(* IEC 61131-3 sources: s7-to-codesys/src/POUs/Lang/Converted/FB_ConveyorStl, 2 files *)

(* ---- FB_ConveyorStl.decl.st ---- *)
// Назначение: Конвейер выдачи реагента (STL, таймеры S5)
//             Ленточный конвейер выдачи реагента (STL S7-300); таймеры T1–T5 и счётчик C1 S5 — глобальные.
//             1. Запрос xReq: S по xStart, затем R по xStop OR xJam (сброс главнее; xJam — прошлого вызова).
//             2. Сирена: SP T1 1 с по фронту xReq, xHorn = T1; снятие запроса обрывает. 3. SD T2 2 с, RLO = xReq.
//             4. Выбег: SF T3 3 с, RLO = T2, xMotor = T3. 5. Поток: SE T4 4 с по фронту xSensor, xFlowOk = T4;
//             взвод SS T5 5 с по фронту xMotor, R T5 при xMotor = 0; затор T5 AND NOT T4 → S xJam; xAck: FR T4
//             (при удерживаемом xSensor контроль запускается снова), R xJam.
//             6. iDelayLeft := L T2 (остаток задержки, единицы 10 мс), wRunOutBcd := LC T3 (BCD со шкалой).
//             7. Счётчик C1: CU по xSensor, R по xCountReset (по уровню); iCount := L C1, wCountBcd := LC C1.
// Автор:      WTP2 (исходный блок S7); перевод в ST — s7conv 0.1.0
// Версия:     0.1 (исходный блок S7)
// Документ:   docs/CONVERSION_REPORT.md, docs/MAPPING.md
// Источник:   samples/lang/FB_ConveyorStl.xml, STL, SW.Blocks.FB "FB_ConveyorStl", пространство имён Interface/v5,
//             FAMILY Dosing
// Сгенерировано s7conv: пометки MIGRATION-CHECK и MIGRATION-TODO требуют ручного разбора.
// MIGRATION-CHECK: стандартный (неоптимизированный) доступ S7: абсолютная адресация и порядок байтов не переносятся
//                  (FB_ConveyorStl.xml, SW.Blocks.FB «FB_ConveyorStl»)
FUNCTION_BLOCK FB_ConveyorStl
VAR_INPUT
    xStart : BOOL;  // Пуск ленты
    xStop : BOOL;  // Стоп ленты
    xSensor : BOOL;  // Датчик изделия на выходе ленты
    xAck : BOOL;  // Квитирование аварии
    xCountReset : BOOL;  // Сброс счётчика изделий
END_VAR
VAR_OUTPUT
    xHorn : BOOL;  // Сирена перед пуском
    xMotor : BOOL;  // Двигатель ленты
    xFlowOk : BOOL;  // Поток изделий в норме (идёт T4)
    xJam : BOOL;  // Авария: затор
    iDelayLeft : INT;  // Остаток задержки пуска, единицы 10 мс
    wRunOutBcd : WORD;  // Остаток выбега, BCD со шкалой
    iCount : INT;  // Изделий
    wCountBcd : WORD;  // Изделий, BCD
END_VAR
VAR
    xReq : BOOL;  // Запрос работы
END_VAR

(* ---- FB_ConveyorStl.impl.st ---- *)
// Сеть 1: Запрос работы
IF xStart THEN
    xReq := TRUE;
END_IF
IF xStop OR xJam THEN
    xReq := FALSE;
END_IF
// Сеть 2: Сирена 1 с при запросе (SP)
// MIGRATION-CHECK: SP T1 → F_S5Pulse (S7Compat): время — F_S7Now(), остаток пересчитывается при обращении к
//                  таймеру; фаза часового процесса CPU (точность ±1 единица шкалы) не моделируется
//                  (FB_ConveyorStl.xml, сеть 2, строка 3)
F_S5Pulse(stTimer := GVL_S5Timers_Lang.aTimer[1], xRlo := xReq, wS5Time := F_S5TimeWord(T#1S));
xHorn := F_S5Q(stTimer := GVL_S5Timers_Lang.aTimer[1]);
// Сеть 3: Задержка пуска 2 с (SD)
// MIGRATION-CHECK: SD T2 → F_S5OnDelay (S7Compat): время — F_S7Now(), остаток пересчитывается при обращении к
//                  таймеру; фаза часового процесса CPU (точность ±1 единица шкалы) не моделируется
//                  (FB_ConveyorStl.xml, сеть 3, строка 3)
F_S5OnDelay(stTimer := GVL_S5Timers_Lang.aTimer[2], xRlo := xReq, wS5Time := F_S5TimeWord(T#2S));
// Сеть 4: Выбег 3 с после снятия запроса (SF)
// MIGRATION-CHECK: SF T3 → F_S5OffDelay (S7Compat): время — F_S7Now(), остаток пересчитывается при обращении к
//                  таймеру; фаза часового процесса CPU (точность ±1 единица шкалы) не моделируется
//                  (FB_ConveyorStl.xml, сеть 4, строка 3)
F_S5OffDelay(stTimer := GVL_S5Timers_Lang.aTimer[3],
             xRlo := F_S5Q(stTimer := GVL_S5Timers_Lang.aTimer[2]),
             wS5Time := F_S5TimeWord(T#3S));
xMotor := F_S5Q(stTimer := GVL_S5Timers_Lang.aTimer[3]);
// Сеть 5: Контроль потока (SE) и затор (SS)
// MIGRATION-CHECK: SE T4 → F_S5ExtPulse (S7Compat): время — F_S7Now(), остаток пересчитывается при обращении к
//                  таймеру; фаза часового процесса CPU (точность ±1 единица шкалы) не моделируется
//                  (FB_ConveyorStl.xml, сеть 5, строка 3)
F_S5ExtPulse(stTimer := GVL_S5Timers_Lang.aTimer[4], xRlo := xSensor, wS5Time := F_S5TimeWord(T#4S));
xFlowOk := F_S5Q(stTimer := GVL_S5Timers_Lang.aTimer[4]);
// MIGRATION-CHECK: SS T5 → F_S5RetOnDelay (S7Compat): время — F_S7Now(), остаток пересчитывается при обращении к
//                  таймеру; фаза часового процесса CPU (точность ±1 единица шкалы) не моделируется
//                  (FB_ConveyorStl.xml, сеть 5, строка 8)
F_S5RetOnDelay(stTimer := GVL_S5Timers_Lang.aTimer[5], xRlo := xMotor, wS5Time := F_S5TimeWord(T#5S));
F_S5Reset(stTimer := GVL_S5Timers_Lang.aTimer[5], xRlo := NOT xMotor);
IF F_S5Q(stTimer := GVL_S5Timers_Lang.aTimer[5]) AND NOT F_S5Q(stTimer := GVL_S5Timers_Lang.aTimer[4]) THEN
    xJam := TRUE;
END_IF
F_S5Enable(stTimer := GVL_S5Timers_Lang.aTimer[4], xRlo := xAck);
IF xAck THEN
    xJam := FALSE;
END_IF
// Сеть 6: Диагностика: остатки таймеров
iDelayLeft := WORD_TO_INT(F_S5Bin(stTimer := GVL_S5Timers_Lang.aTimer[2]));
wRunOutBcd := F_S5Bcd(stTimer := GVL_S5Timers_Lang.aTimer[3]);
// Сеть 7: Счётчик изделий (C1)
F_S5CountUp(stCounter := GVL_S5Counters_Lang.aCounter[1], xRlo := xSensor);
F_S5CounterReset(stCounter := GVL_S5Counters_Lang.aCounter[1], xRlo := xCountReset);
iCount := WORD_TO_INT(F_S5CounterBin(stCounter := GVL_S5Counters_Lang.aCounter[1]));
wCountBcd := F_S5CounterBcd(stCounter := GVL_S5Counters_Lang.aCounter[1]);
